// TIA Portal V20 export
FUNCTION_BLOCK "PR_MultiPosShuttle_Soft2.0 1_workflow_268c4d"   // FB49, LAD
{ S7_Optimized_Access := 'TRUE' }
// stored: MemoryReserve 100, SetENOAutomatically false
   VAR_INPUT
      iAutoRunning : Bool;
      iFaultReset : Bool;
      iGantry2Safe : Bool;
      iGantry_2Safe : Bool;
      iHIPOTTesSafe : Bool;
      iHIPOTTestOver : Bool;
      iHipotTestSafe : Bool;
      iInfeedGantrySafe : Bool;
      iOTS_Frm_Gantry : Bool;
      iPartPresent : Bool;
      iPartPrsent : Bool;
      iRTR_Frm_Gantry2 : Bool;
      iReset_fault : Bool;
      iShuttleAtGantry2Pos : Bool;
      iShuttleAtGantry_2Pos : Bool;
      iShuttleAtHIPOTPos : Bool;
      iShuttleAtHIPOTTestPos : Bool;
      iShuttleAtPartLoadPos : Bool;
      iSstMode : Bool;
      iSstPB : Bool;
   END_VAR
   VAR_OUTPUT
      qError : Array[0..10] of Bool;
      qHiPotTestStartCmd : Bool;
      qMessage : Array[0..10] of Bool;
      qRTR_To_InfeedGantry : Bool;
      qShuttleGantry_2PosCmd : Bool;
      qShuttleHIPOTTestPosCmd : Bool;
      qStateNo : Int;
      qShuttleReceivePosCmd : Bool;
   END_VAR
   VAR
      c10_ChkRecCond_T1 : Bool;
      c10_ChkRecCond_T2 : Bool;
      c10_ChkRecCond_T3 : Bool;
      c10_ChkRecCond_T4 : Bool;
      c10_ChkRecCond_T5 : Bool;
      c150_ChkOprnSts_T1 : Bool;
      c150_ChkOprnSts_T2 : Bool;
      c30_ChkPartPrsnt_T1 : Bool;
      c30_ChkPartPrsnt_T2 : Bool;
      s100_WtHipotTestOver : Bool;
      s100_WtHipotTestOver_T1 : Bool;
      s10_ChkRecCond : Bool;
      s10_ChkRecCond_T1 : Bool;
      s10_ChkRecCond_T2 : Bool;
      s10_ChkRecCond_T3 : Bool;
      s10_ChkRecCond_T4 : Bool;
      s10_ChkRecCond_T5 : Bool;
      s110_WtGantry2Safe : Bool;
      s110_WtGantry2Safe_T1 : Bool;
      s120_WtShtlGantry2Pos : Bool;
      s120_WtShtlGantry2Pos_T1 : Bool;
      s130_WtRTRFrmGantry2 : Bool;
      s130_WtRTRFrmGantry2_T1 : Bool;
      s140_WtPartAbsntGantry2Safe : Bool;
      s140_WtPartAbsntGantry2Safe_T1 : Bool;
      s150_ChkOprnSts : Bool;
      s150_ChkOprnSts_T1 : Bool;
      s150_ChkOprnSts_T2 : Bool;
      s1_WtResetRel : Bool;
      s1_WtResetRel_T1 : Bool;
      s20_WtFaultReset : Bool;
      s20_WtFaultReset_T1 : Bool;
      s30_ChkPartPrsnt : Bool;
      s30_ChkPartPrsnt_T1 : Bool;
      s30_ChkPartPrsnt_T2 : Bool;
      s40_WtAllSysSafe : Bool;
      s40_WtAllSysSafe_T1 : Bool;
      s50_WtShtlPartRcvPos : Bool;
      s50_WtShtlPartRcvPos_T1 : Bool;
      s60_WtOTSFrmGantry : Bool;
      s60_WtOTSFrmGantry_T1 : Bool;
      s70_WtPartPlcdGantrySafe : Bool;
      s70_WtPartPlcdGantrySafe_T1 : Bool;
      s80_WtHIPOTSafe : Bool;
      s80_WtHIPOTSafe_T1 : Bool;
      s90_WtShtlHIPOTPos : Bool;
      s90_WtShtlHIPOTPos_T1 : Bool;
      sHIPOTOprnOver : Bool;
      sHipotTestInProgress : Bool;
      sPickInProgress : Bool;
      sPlaceInProgress : Bool;
      sSst : Bool;
      sSstPulse : Bool;
      sSstRise : Bool;
      sStWtResetRel : Bool;
      sStWtResetRel_T1 : Bool;
   END_VAR
   VAR_TEMP
      tOne : Bool;
   END_VAR
   VAR_TEMP   // added for the SCL form of the ladder/FBD networks
      _w1 : Bool;
      _w2 : Bool;
      _w3 : Bool;
      _w4 : Bool;
   END_VAR
BEGIN

REGION Network 1
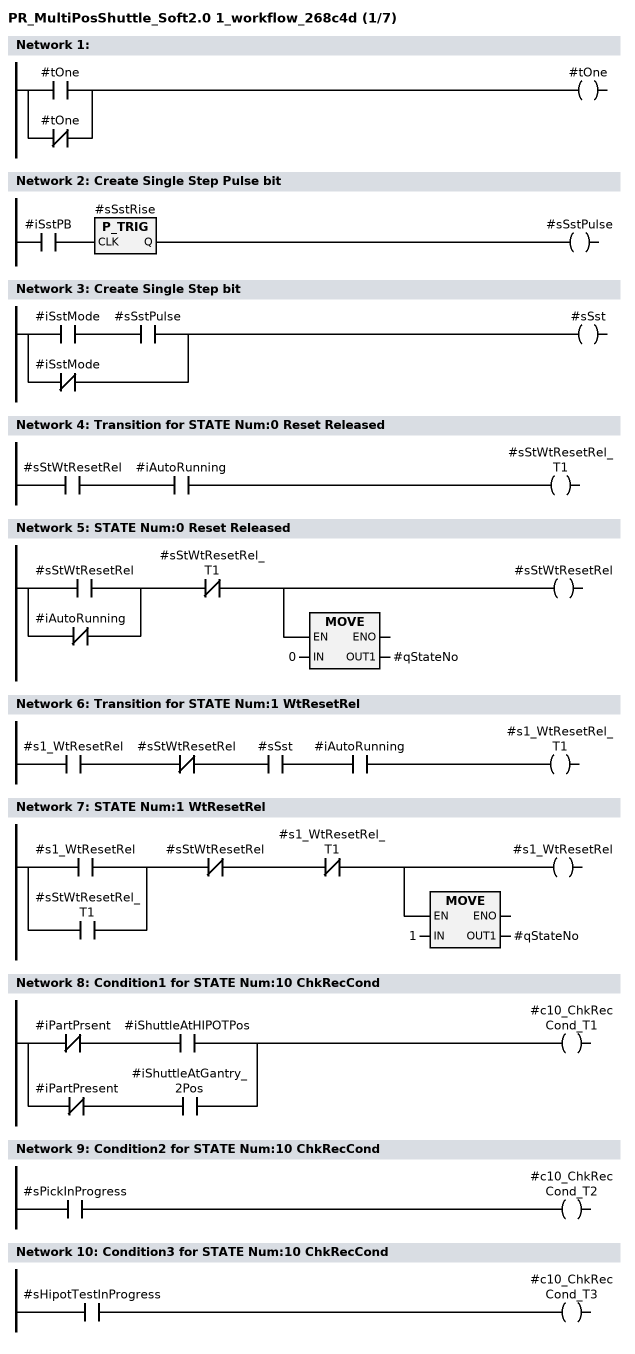
   RUNG wire#powerrail
      Contact( #tOne )
      wire#w1
      Coil( #tOne )
   END_RUNG
   RUNG wire#powerrail
      I_Contact( #tOne )
   END_RUNG wire#w1
   // the same network as SCL:
   #tOne := #tOne OR NOT #tOne;
END_REGION

REGION Network 2: Create Single Step Pulse bit
   RUNG wire#powerrail
      Contact( #iSstPB )
      P_Trig( #sSstRise )
      Coil( #sSstPulse )
   END_RUNG
   // the same network as SCL:
   #_w1 := #iSstPB AND NOT #sSstRise;   // rising edge
   #sSstRise := #iSstPB;
   #sSstPulse := #_w1;
END_REGION

REGION Network 3: Create Single Step bit
   RUNG wire#powerrail
      Contact( #iSstMode )
      Contact( #sSstPulse )
      wire#w1
      Coil( #sSst )
   END_RUNG
   RUNG wire#powerrail
      I_Contact( #iSstMode )
   END_RUNG wire#w1
   // the same network as SCL:
   #sSst := (#iSstMode AND #sSstPulse) OR NOT #iSstMode;
END_REGION

REGION Network 4: Transition for STATE Num:0 Reset Released
   RUNG wire#powerrail
      Contact( #sStWtResetRel )
      Contact( #iAutoRunning )
      Coil( #sStWtResetRel_T1 )
   END_RUNG
   // the same network as SCL:
   #sStWtResetRel_T1 := #sStWtResetRel AND #iAutoRunning;
END_REGION

REGION Network 5: STATE Num:0 Reset Released
   RUNG wire#powerrail
      Contact( #sStWtResetRel )
      wire#w1
      I_Contact( #sStWtResetRel_T1 )
      wire#w2
      Coil( #sStWtResetRel )
   END_RUNG
   RUNG wire#powerrail
      I_Contact( #iAutoRunning )
   END_RUNG wire#w1
   RUNG wire#w2
      { S7_GenerateENO := "TRUE" } Move(in := 0, out1 => #qStateNo)
   END_RUNG
   // the same network as SCL:
   #sStWtResetRel := (#sStWtResetRel OR NOT #iAutoRunning) AND NOT #sStWtResetRel_T1;
   IF #sStWtResetRel THEN #qStateNo := 0; END_IF;
END_REGION

REGION Network 6: Transition for STATE Num:1 WtResetRel
   RUNG wire#powerrail
      Contact( #s1_WtResetRel )
      I_Contact( #sStWtResetRel )
      Contact( #sSst )
      Contact( #iAutoRunning )
      Coil( #s1_WtResetRel_T1 )
   END_RUNG
   // the same network as SCL:
   #s1_WtResetRel_T1 := #s1_WtResetRel AND NOT #sStWtResetRel AND #sSst AND #iAutoRunning;
END_REGION

REGION Network 7: STATE Num:1 WtResetRel
   RUNG wire#powerrail
      Contact( #s1_WtResetRel )
      wire#w1
      I_Contact( #sStWtResetRel )
      I_Contact( #s1_WtResetRel_T1 )
      wire#w2
      Coil( #s1_WtResetRel )
   END_RUNG
   RUNG wire#powerrail
      Contact( #sStWtResetRel_T1 )
   END_RUNG wire#w1
   RUNG wire#w2
      { S7_GenerateENO := "TRUE" } Move(in := 1, out1 => #qStateNo)
   END_RUNG
   // the same network as SCL:
   #s1_WtResetRel := (#s1_WtResetRel OR #sStWtResetRel_T1) AND NOT #sStWtResetRel AND NOT #s1_WtResetRel_T1;
   IF #s1_WtResetRel THEN #qStateNo := 1; END_IF;
END_REGION

REGION Network 8: Condition1 for STATE Num:10 ChkRecCond
   RUNG wire#powerrail
      I_Contact( #iPartPrsent )
      Contact( #iShuttleAtHIPOTPos )
      wire#w1
      Coil( #c10_ChkRecCond_T1 )
   END_RUNG
   RUNG wire#powerrail
      I_Contact( #iPartPresent )
      Contact( #iShuttleAtGantry_2Pos )
   END_RUNG wire#w1
   // the same network as SCL:
   #c10_ChkRecCond_T1 := (NOT #iPartPrsent AND #iShuttleAtHIPOTPos) OR (NOT #iPartPresent AND #iShuttleAtGantry_2Pos);
END_REGION

REGION Network 9: Condition2 for STATE Num:10 ChkRecCond
   RUNG wire#powerrail
      Contact( #sPickInProgress )
      Coil( #c10_ChkRecCond_T2 )
   END_RUNG
   // the same network as SCL:
   #c10_ChkRecCond_T2 := #sPickInProgress;
END_REGION

REGION Network 10: Condition3 for STATE Num:10 ChkRecCond
   RUNG wire#powerrail
      Contact( #sHipotTestInProgress )
      Coil( #c10_ChkRecCond_T3 )
   END_RUNG
   // the same network as SCL:
   #c10_ChkRecCond_T3 := #sHipotTestInProgress;
END_REGION

REGION Network 11: Condition4 for STATE Num:10 ChkRecCond
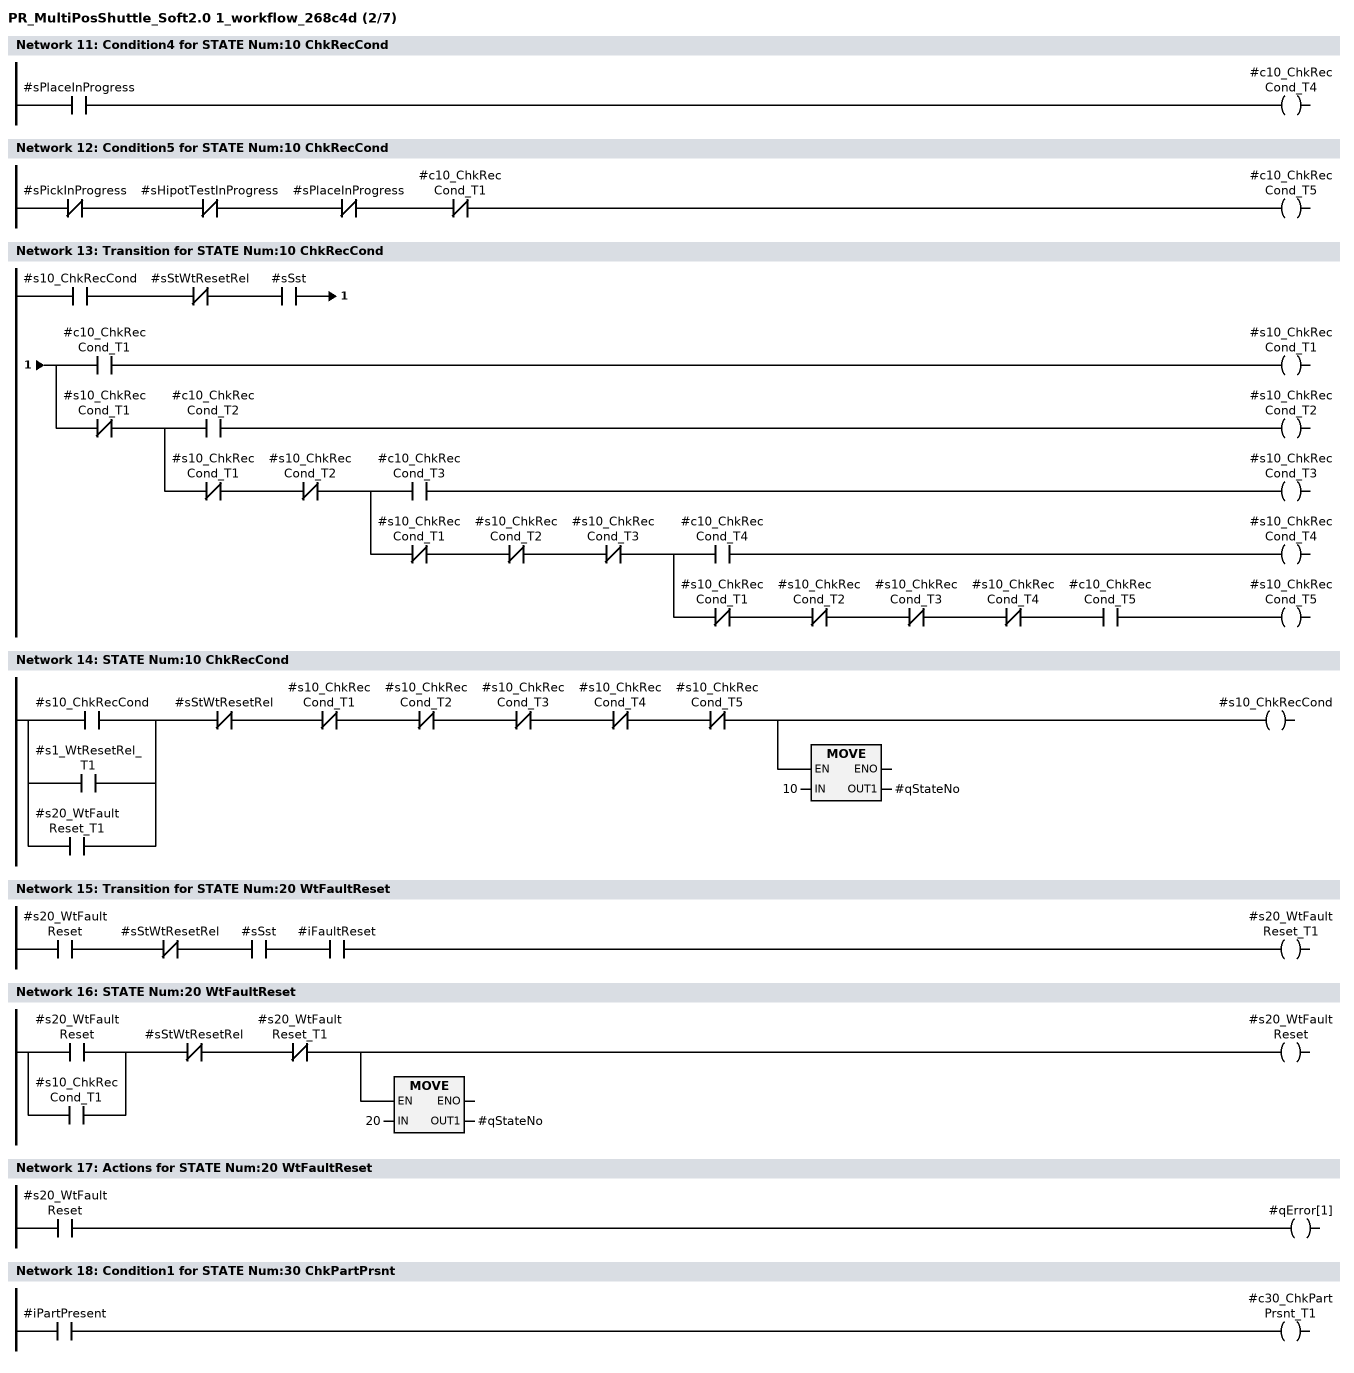
   RUNG wire#powerrail
      Contact( #sPlaceInProgress )
      Coil( #c10_ChkRecCond_T4 )
   END_RUNG
   // the same network as SCL:
   #c10_ChkRecCond_T4 := #sPlaceInProgress;
END_REGION

REGION Network 12: Condition5 for STATE Num:10 ChkRecCond
   RUNG wire#powerrail
      I_Contact( #sPickInProgress )
      I_Contact( #sHipotTestInProgress )
      I_Contact( #sPlaceInProgress )
      I_Contact( #c10_ChkRecCond_T1 )
      Coil( #c10_ChkRecCond_T5 )
   END_RUNG
   // the same network as SCL:
   #c10_ChkRecCond_T5 := NOT #sPickInProgress AND NOT #sHipotTestInProgress AND NOT #sPlaceInProgress AND NOT #c10_ChkRecCond_T1;
END_REGION

REGION Network 13: Transition for STATE Num:10 ChkRecCond
   RUNG wire#powerrail
      Contact( #s10_ChkRecCond )
      I_Contact( #sStWtResetRel )
      Contact( #sSst )
      wire#w1
      Contact( #c10_ChkRecCond_T1 )
      Coil( #s10_ChkRecCond_T1 )
   END_RUNG
   RUNG wire#w1
      I_Contact( #s10_ChkRecCond_T1 )
      wire#w2
      Contact( #c10_ChkRecCond_T2 )
      Coil( #s10_ChkRecCond_T2 )
   END_RUNG
   RUNG wire#w2
      I_Contact( #s10_ChkRecCond_T1 )
      I_Contact( #s10_ChkRecCond_T2 )
      wire#w3
      Contact( #c10_ChkRecCond_T3 )
      Coil( #s10_ChkRecCond_T3 )
   END_RUNG
   RUNG wire#w3
      I_Contact( #s10_ChkRecCond_T1 )
      I_Contact( #s10_ChkRecCond_T2 )
      I_Contact( #s10_ChkRecCond_T3 )
      wire#w4
      Contact( #c10_ChkRecCond_T4 )
      Coil( #s10_ChkRecCond_T4 )
   END_RUNG
   RUNG wire#w4
      I_Contact( #s10_ChkRecCond_T1 )
      I_Contact( #s10_ChkRecCond_T2 )
      I_Contact( #s10_ChkRecCond_T3 )
      I_Contact( #s10_ChkRecCond_T4 )
      Contact( #c10_ChkRecCond_T5 )
      Coil( #s10_ChkRecCond_T5 )
   END_RUNG
   // the same network as SCL:
   #_w1 := #s10_ChkRecCond AND NOT #sStWtResetRel AND #sSst;
   #s10_ChkRecCond_T1 := #_w1 AND #c10_ChkRecCond_T1;
   #_w2 := #_w1 AND NOT #s10_ChkRecCond_T1;
   #s10_ChkRecCond_T2 := #_w2 AND #c10_ChkRecCond_T2;
   #_w3 := #_w2 AND NOT #s10_ChkRecCond_T1 AND NOT #s10_ChkRecCond_T2;
   #s10_ChkRecCond_T3 := #_w3 AND #c10_ChkRecCond_T3;
   #_w4 := #_w3 AND NOT #s10_ChkRecCond_T1 AND NOT #s10_ChkRecCond_T2 AND NOT #s10_ChkRecCond_T3;
   #s10_ChkRecCond_T4 := #_w4 AND #c10_ChkRecCond_T4;
   #s10_ChkRecCond_T5 := #_w4 AND NOT #s10_ChkRecCond_T1 AND NOT #s10_ChkRecCond_T2 AND NOT #s10_ChkRecCond_T3 AND NOT #s10_ChkRecCond_T4 AND #c10_ChkRecCond_T5;
END_REGION

REGION Network 14: STATE Num:10 ChkRecCond
   RUNG wire#powerrail
      Contact( #s10_ChkRecCond )
      wire#w1
      I_Contact( #sStWtResetRel )
      I_Contact( #s10_ChkRecCond_T1 )
      I_Contact( #s10_ChkRecCond_T2 )
      I_Contact( #s10_ChkRecCond_T3 )
      I_Contact( #s10_ChkRecCond_T4 )
      I_Contact( #s10_ChkRecCond_T5 )
      wire#w2
      Coil( #s10_ChkRecCond )
   END_RUNG
   RUNG wire#powerrail
      Contact( #s1_WtResetRel_T1 )
   END_RUNG wire#w1
   RUNG wire#powerrail
      Contact( #s20_WtFaultReset_T1 )
   END_RUNG wire#w1
   RUNG wire#w2
      { S7_GenerateENO := "TRUE" } Move(in := 10, out1 => #qStateNo)
   END_RUNG
   // the same network as SCL:
   #s10_ChkRecCond := (#s10_ChkRecCond OR #s1_WtResetRel_T1 OR #s20_WtFaultReset_T1) AND NOT #sStWtResetRel AND NOT #s10_ChkRecCond_T1 AND NOT #s10_ChkRecCond_T2 AND NOT #s10_ChkRecCond_T3 AND NOT #s10_ChkRecCond_T4 AND NOT #s10_ChkRecCond_T5;
   IF #s10_ChkRecCond THEN #qStateNo := 10; END_IF;
END_REGION

REGION Network 15: Transition for STATE Num:20 WtFaultReset
   RUNG wire#powerrail
      Contact( #s20_WtFaultReset )
      I_Contact( #sStWtResetRel )
      Contact( #sSst )
      Contact( #iFaultReset )
      Coil( #s20_WtFaultReset_T1 )
   END_RUNG
   // the same network as SCL:
   #s20_WtFaultReset_T1 := #s20_WtFaultReset AND NOT #sStWtResetRel AND #sSst AND #iFaultReset;
END_REGION

REGION Network 16: STATE Num:20 WtFaultReset
   RUNG wire#powerrail
      Contact( #s20_WtFaultReset )
      wire#w1
      I_Contact( #sStWtResetRel )
      I_Contact( #s20_WtFaultReset_T1 )
      wire#w2
      Coil( #s20_WtFaultReset )
   END_RUNG
   RUNG wire#powerrail
      Contact( #s10_ChkRecCond_T1 )
   END_RUNG wire#w1
   RUNG wire#w2
      { S7_GenerateENO := "TRUE" } Move(in := 20, out1 => #qStateNo)
   END_RUNG
   // the same network as SCL:
   #s20_WtFaultReset := (#s20_WtFaultReset OR #s10_ChkRecCond_T1) AND NOT #sStWtResetRel AND NOT #s20_WtFaultReset_T1;
   IF #s20_WtFaultReset THEN #qStateNo := 20; END_IF;
END_REGION

REGION Network 17: Actions for STATE Num:20 WtFaultReset
   RUNG wire#powerrail
      Contact( #s20_WtFaultReset )
      Coil( #qError[1] )
   END_RUNG
   // the same network as SCL:
   #qError[1] := #s20_WtFaultReset;
END_REGION

REGION Network 18: Condition1 for STATE Num:30 ChkPartPrsnt
   RUNG wire#powerrail
      Contact( #iPartPresent )
      Coil( #c30_ChkPartPrsnt_T1 )
   END_RUNG
   // the same network as SCL:
   #c30_ChkPartPrsnt_T1 := #iPartPresent;
END_REGION

REGION Network 19: Condition2 for STATE Num:30 ChkPartPrsnt
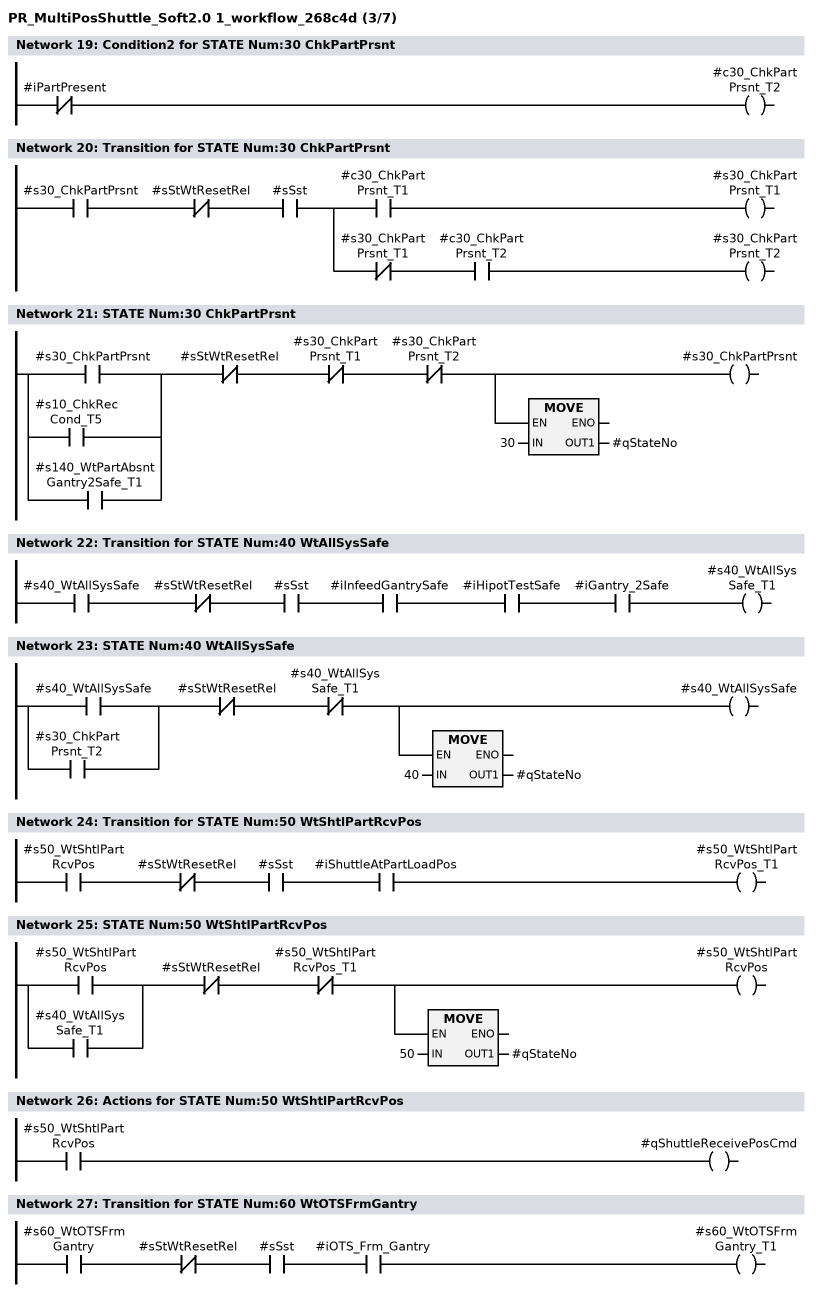
   RUNG wire#powerrail
      I_Contact( #iPartPresent )
      Coil( #c30_ChkPartPrsnt_T2 )
   END_RUNG
   // the same network as SCL:
   #c30_ChkPartPrsnt_T2 := NOT #iPartPresent;
END_REGION

REGION Network 20: Transition for STATE Num:30 ChkPartPrsnt
   RUNG wire#powerrail
      Contact( #s30_ChkPartPrsnt )
      I_Contact( #sStWtResetRel )
      Contact( #sSst )
      wire#w1
      Contact( #c30_ChkPartPrsnt_T1 )
      Coil( #s30_ChkPartPrsnt_T1 )
   END_RUNG
   RUNG wire#w1
      I_Contact( #s30_ChkPartPrsnt_T1 )
      Contact( #c30_ChkPartPrsnt_T2 )
      Coil( #s30_ChkPartPrsnt_T2 )
   END_RUNG
   // the same network as SCL:
   #_w1 := #s30_ChkPartPrsnt AND NOT #sStWtResetRel AND #sSst;
   #s30_ChkPartPrsnt_T1 := #_w1 AND #c30_ChkPartPrsnt_T1;
   #s30_ChkPartPrsnt_T2 := #_w1 AND NOT #s30_ChkPartPrsnt_T1 AND #c30_ChkPartPrsnt_T2;
END_REGION

REGION Network 21: STATE Num:30 ChkPartPrsnt
   RUNG wire#powerrail
      Contact( #s30_ChkPartPrsnt )
      wire#w1
      I_Contact( #sStWtResetRel )
      I_Contact( #s30_ChkPartPrsnt_T1 )
      I_Contact( #s30_ChkPartPrsnt_T2 )
      wire#w2
      Coil( #s30_ChkPartPrsnt )
   END_RUNG
   RUNG wire#powerrail
      Contact( #s10_ChkRecCond_T5 )
   END_RUNG wire#w1
   RUNG wire#powerrail
      Contact( #s140_WtPartAbsntGantry2Safe_T1 )
   END_RUNG wire#w1
   RUNG wire#w2
      { S7_GenerateENO := "TRUE" } Move(in := 30, out1 => #qStateNo)
   END_RUNG
   // the same network as SCL:
   #s30_ChkPartPrsnt := (#s30_ChkPartPrsnt OR #s10_ChkRecCond_T5 OR #s140_WtPartAbsntGantry2Safe_T1) AND NOT #sStWtResetRel AND NOT #s30_ChkPartPrsnt_T1 AND NOT #s30_ChkPartPrsnt_T2;
   IF #s30_ChkPartPrsnt THEN #qStateNo := 30; END_IF;
END_REGION

REGION Network 22: Transition for STATE Num:40 WtAllSysSafe
   RUNG wire#powerrail
      Contact( #s40_WtAllSysSafe )
      I_Contact( #sStWtResetRel )
      Contact( #sSst )
      Contact( #iInfeedGantrySafe )
      Contact( #iHipotTestSafe )
      Contact( #iGantry_2Safe )
      Coil( #s40_WtAllSysSafe_T1 )
   END_RUNG
   // the same network as SCL:
   #s40_WtAllSysSafe_T1 := #s40_WtAllSysSafe AND NOT #sStWtResetRel AND #sSst AND #iInfeedGantrySafe AND #iHipotTestSafe AND #iGantry_2Safe;
END_REGION

REGION Network 23: STATE Num:40 WtAllSysSafe
   RUNG wire#powerrail
      Contact( #s40_WtAllSysSafe )
      wire#w1
      I_Contact( #sStWtResetRel )
      I_Contact( #s40_WtAllSysSafe_T1 )
      wire#w2
      Coil( #s40_WtAllSysSafe )
   END_RUNG
   RUNG wire#powerrail
      Contact( #s30_ChkPartPrsnt_T2 )
   END_RUNG wire#w1
   RUNG wire#w2
      { S7_GenerateENO := "TRUE" } Move(in := 40, out1 => #qStateNo)
   END_RUNG
   // the same network as SCL:
   #s40_WtAllSysSafe := (#s40_WtAllSysSafe OR #s30_ChkPartPrsnt_T2) AND NOT #sStWtResetRel AND NOT #s40_WtAllSysSafe_T1;
   IF #s40_WtAllSysSafe THEN #qStateNo := 40; END_IF;
END_REGION

REGION Network 24: Transition for STATE Num:50 WtShtlPartRcvPos
   RUNG wire#powerrail
      Contact( #s50_WtShtlPartRcvPos )
      I_Contact( #sStWtResetRel )
      Contact( #sSst )
      Contact( #iShuttleAtPartLoadPos )
      Coil( #s50_WtShtlPartRcvPos_T1 )
   END_RUNG
   // the same network as SCL:
   #s50_WtShtlPartRcvPos_T1 := #s50_WtShtlPartRcvPos AND NOT #sStWtResetRel AND #sSst AND #iShuttleAtPartLoadPos;
END_REGION

REGION Network 25: STATE Num:50 WtShtlPartRcvPos
   RUNG wire#powerrail
      Contact( #s50_WtShtlPartRcvPos )
      wire#w1
      I_Contact( #sStWtResetRel )
      I_Contact( #s50_WtShtlPartRcvPos_T1 )
      wire#w2
      Coil( #s50_WtShtlPartRcvPos )
   END_RUNG
   RUNG wire#powerrail
      Contact( #s40_WtAllSysSafe_T1 )
   END_RUNG wire#w1
   RUNG wire#w2
      { S7_GenerateENO := "TRUE" } Move(in := 50, out1 => #qStateNo)
   END_RUNG
   // the same network as SCL:
   #s50_WtShtlPartRcvPos := (#s50_WtShtlPartRcvPos OR #s40_WtAllSysSafe_T1) AND NOT #sStWtResetRel AND NOT #s50_WtShtlPartRcvPos_T1;
   IF #s50_WtShtlPartRcvPos THEN #qStateNo := 50; END_IF;
END_REGION

REGION Network 26: Actions for STATE Num:50 WtShtlPartRcvPos
   RUNG wire#powerrail
      Contact( #s50_WtShtlPartRcvPos )
      Coil( #qShuttleReceivePosCmd )
   END_RUNG
   // the same network as SCL:
   #qShuttleReceivePosCmd := #s50_WtShtlPartRcvPos;
END_REGION

REGION Network 27: Transition for STATE Num:60 WtOTSFrmGantry
   RUNG wire#powerrail
      Contact( #s60_WtOTSFrmGantry )
      I_Contact( #sStWtResetRel )
      Contact( #sSst )
      Contact( #iOTS_Frm_Gantry )
      Coil( #s60_WtOTSFrmGantry_T1 )
   END_RUNG
   // the same network as SCL:
   #s60_WtOTSFrmGantry_T1 := #s60_WtOTSFrmGantry AND NOT #sStWtResetRel AND #sSst AND #iOTS_Frm_Gantry;
END_REGION

REGION Network 28: STATE Num:60 WtOTSFrmGantry
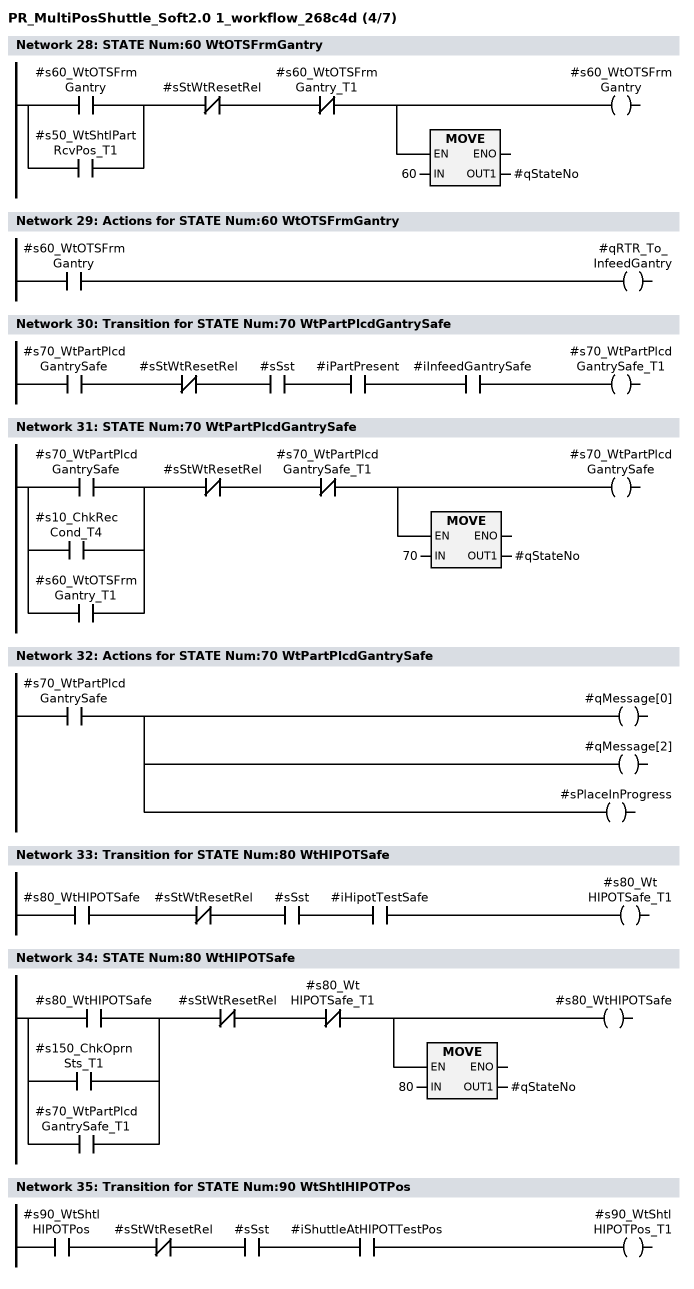
   RUNG wire#powerrail
      Contact( #s60_WtOTSFrmGantry )
      wire#w1
      I_Contact( #sStWtResetRel )
      I_Contact( #s60_WtOTSFrmGantry_T1 )
      wire#w2
      Coil( #s60_WtOTSFrmGantry )
   END_RUNG
   RUNG wire#powerrail
      Contact( #s50_WtShtlPartRcvPos_T1 )
   END_RUNG wire#w1
   RUNG wire#w2
      { S7_GenerateENO := "TRUE" } Move(in := 60, out1 => #qStateNo)
   END_RUNG
   // the same network as SCL:
   #s60_WtOTSFrmGantry := (#s60_WtOTSFrmGantry OR #s50_WtShtlPartRcvPos_T1) AND NOT #sStWtResetRel AND NOT #s60_WtOTSFrmGantry_T1;
   IF #s60_WtOTSFrmGantry THEN #qStateNo := 60; END_IF;
END_REGION

REGION Network 29: Actions for STATE Num:60 WtOTSFrmGantry
   RUNG wire#powerrail
      Contact( #s60_WtOTSFrmGantry )
      Coil( #qRTR_To_InfeedGantry )
   END_RUNG
   // the same network as SCL:
   #qRTR_To_InfeedGantry := #s60_WtOTSFrmGantry;
END_REGION

REGION Network 30: Transition for STATE Num:70 WtPartPlcdGantrySafe
   RUNG wire#powerrail
      Contact( #s70_WtPartPlcdGantrySafe )
      I_Contact( #sStWtResetRel )
      Contact( #sSst )
      Contact( #iPartPresent )
      Contact( #iInfeedGantrySafe )
      Coil( #s70_WtPartPlcdGantrySafe_T1 )
   END_RUNG
   // the same network as SCL:
   #s70_WtPartPlcdGantrySafe_T1 := #s70_WtPartPlcdGantrySafe AND NOT #sStWtResetRel AND #sSst AND #iPartPresent AND #iInfeedGantrySafe;
END_REGION

REGION Network 31: STATE Num:70 WtPartPlcdGantrySafe
   RUNG wire#powerrail
      Contact( #s70_WtPartPlcdGantrySafe )
      wire#w1
      I_Contact( #sStWtResetRel )
      I_Contact( #s70_WtPartPlcdGantrySafe_T1 )
      wire#w2
      Coil( #s70_WtPartPlcdGantrySafe )
   END_RUNG
   RUNG wire#powerrail
      Contact( #s10_ChkRecCond_T4 )
   END_RUNG wire#w1
   RUNG wire#powerrail
      Contact( #s60_WtOTSFrmGantry_T1 )
   END_RUNG wire#w1
   RUNG wire#w2
      { S7_GenerateENO := "TRUE" } Move(in := 70, out1 => #qStateNo)
   END_RUNG
   // the same network as SCL:
   #s70_WtPartPlcdGantrySafe := (#s70_WtPartPlcdGantrySafe OR #s10_ChkRecCond_T4 OR #s60_WtOTSFrmGantry_T1) AND NOT #sStWtResetRel AND NOT #s70_WtPartPlcdGantrySafe_T1;
   IF #s70_WtPartPlcdGantrySafe THEN #qStateNo := 70; END_IF;
END_REGION

REGION Network 32: Actions for STATE Num:70 WtPartPlcdGantrySafe
   RUNG wire#powerrail
      Contact( #s70_WtPartPlcdGantrySafe )
      wire#w1
      Coil( #qMessage[0] )
   END_RUNG
   RUNG wire#w1
      Coil( #qMessage[2] )
   END_RUNG
   RUNG wire#w1
      Coil( #sPlaceInProgress )
   END_RUNG
   // the same network as SCL:
   #qMessage[0] := #s70_WtPartPlcdGantrySafe;
   #qMessage[2] := #s70_WtPartPlcdGantrySafe;
   #sPlaceInProgress := #s70_WtPartPlcdGantrySafe;
END_REGION

REGION Network 33: Transition for STATE Num:80 WtHIPOTSafe
   RUNG wire#powerrail
      Contact( #s80_WtHIPOTSafe )
      I_Contact( #sStWtResetRel )
      Contact( #sSst )
      Contact( #iHipotTestSafe )
      Coil( #s80_WtHIPOTSafe_T1 )
   END_RUNG
   // the same network as SCL:
   #s80_WtHIPOTSafe_T1 := #s80_WtHIPOTSafe AND NOT #sStWtResetRel AND #sSst AND #iHipotTestSafe;
END_REGION

REGION Network 34: STATE Num:80 WtHIPOTSafe
   RUNG wire#powerrail
      Contact( #s80_WtHIPOTSafe )
      wire#w1
      I_Contact( #sStWtResetRel )
      I_Contact( #s80_WtHIPOTSafe_T1 )
      wire#w2
      Coil( #s80_WtHIPOTSafe )
   END_RUNG
   RUNG wire#powerrail
      Contact( #s150_ChkOprnSts_T1 )
   END_RUNG wire#w1
   RUNG wire#powerrail
      Contact( #s70_WtPartPlcdGantrySafe_T1 )
   END_RUNG wire#w1
   RUNG wire#w2
      { S7_GenerateENO := "TRUE" } Move(in := 80, out1 => #qStateNo)
   END_RUNG
   // the same network as SCL:
   #s80_WtHIPOTSafe := (#s80_WtHIPOTSafe OR #s150_ChkOprnSts_T1 OR #s70_WtPartPlcdGantrySafe_T1) AND NOT #sStWtResetRel AND NOT #s80_WtHIPOTSafe_T1;
   IF #s80_WtHIPOTSafe THEN #qStateNo := 80; END_IF;
END_REGION

REGION Network 35: Transition for STATE Num:90 WtShtlHIPOTPos
   RUNG wire#powerrail
      Contact( #s90_WtShtlHIPOTPos )
      I_Contact( #sStWtResetRel )
      Contact( #sSst )
      Contact( #iShuttleAtHIPOTTestPos )
      Coil( #s90_WtShtlHIPOTPos_T1 )
   END_RUNG
   // the same network as SCL:
   #s90_WtShtlHIPOTPos_T1 := #s90_WtShtlHIPOTPos AND NOT #sStWtResetRel AND #sSst AND #iShuttleAtHIPOTTestPos;
END_REGION

REGION Network 36: STATE Num:90 WtShtlHIPOTPos
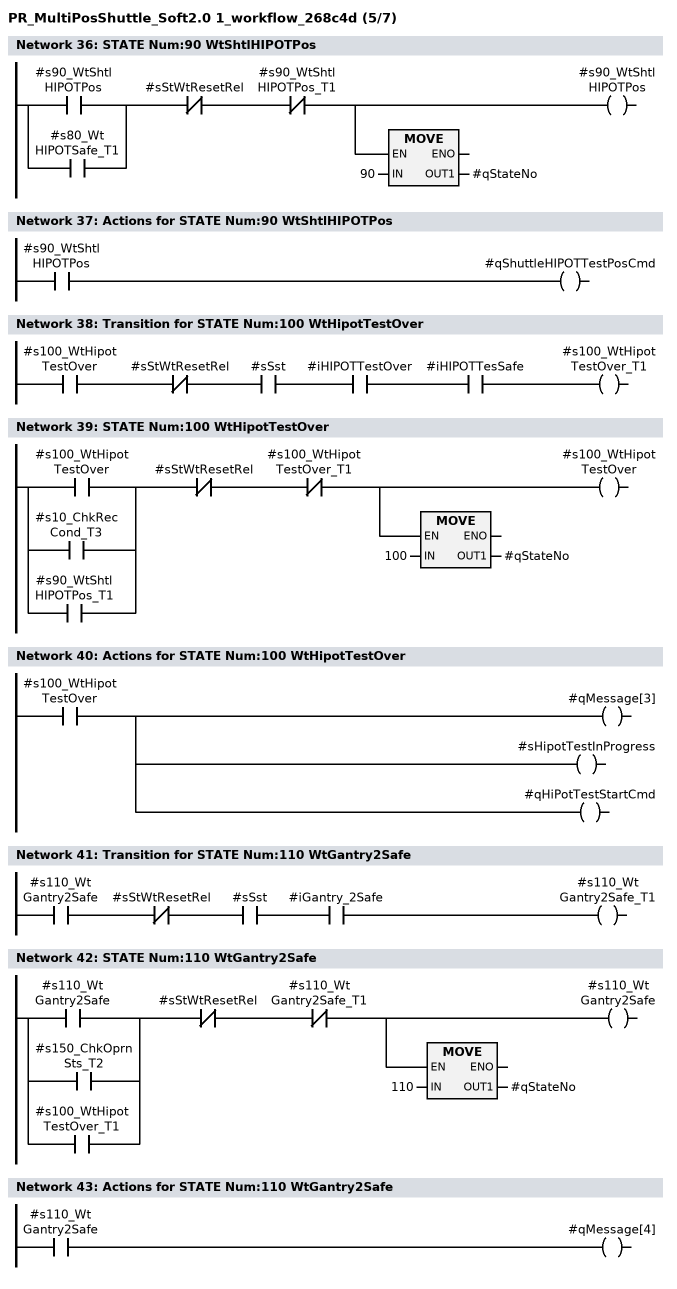
   RUNG wire#powerrail
      Contact( #s90_WtShtlHIPOTPos )
      wire#w1
      I_Contact( #sStWtResetRel )
      I_Contact( #s90_WtShtlHIPOTPos_T1 )
      wire#w2
      Coil( #s90_WtShtlHIPOTPos )
   END_RUNG
   RUNG wire#powerrail
      Contact( #s80_WtHIPOTSafe_T1 )
   END_RUNG wire#w1
   RUNG wire#w2
      { S7_GenerateENO := "TRUE" } Move(in := 90, out1 => #qStateNo)
   END_RUNG
   // the same network as SCL:
   #s90_WtShtlHIPOTPos := (#s90_WtShtlHIPOTPos OR #s80_WtHIPOTSafe_T1) AND NOT #sStWtResetRel AND NOT #s90_WtShtlHIPOTPos_T1;
   IF #s90_WtShtlHIPOTPos THEN #qStateNo := 90; END_IF;
END_REGION

REGION Network 37: Actions for STATE Num:90 WtShtlHIPOTPos
   RUNG wire#powerrail
      Contact( #s90_WtShtlHIPOTPos )
      Coil( #qShuttleHIPOTTestPosCmd )
   END_RUNG
   // the same network as SCL:
   #qShuttleHIPOTTestPosCmd := #s90_WtShtlHIPOTPos;
END_REGION

REGION Network 38: Transition for STATE Num:100 WtHipotTestOver
   RUNG wire#powerrail
      Contact( #s100_WtHipotTestOver )
      I_Contact( #sStWtResetRel )
      Contact( #sSst )
      Contact( #iHIPOTTestOver )
      Contact( #iHIPOTTesSafe )
      Coil( #s100_WtHipotTestOver_T1 )
   END_RUNG
   // the same network as SCL:
   #s100_WtHipotTestOver_T1 := #s100_WtHipotTestOver AND NOT #sStWtResetRel AND #sSst AND #iHIPOTTestOver AND #iHIPOTTesSafe;
END_REGION

REGION Network 39: STATE Num:100 WtHipotTestOver
   RUNG wire#powerrail
      Contact( #s100_WtHipotTestOver )
      wire#w1
      I_Contact( #sStWtResetRel )
      I_Contact( #s100_WtHipotTestOver_T1 )
      wire#w2
      Coil( #s100_WtHipotTestOver )
   END_RUNG
   RUNG wire#powerrail
      Contact( #s10_ChkRecCond_T3 )
   END_RUNG wire#w1
   RUNG wire#powerrail
      Contact( #s90_WtShtlHIPOTPos_T1 )
   END_RUNG wire#w1
   RUNG wire#w2
      { S7_GenerateENO := "TRUE" } Move(in := 100, out1 => #qStateNo)
   END_RUNG
   // the same network as SCL:
   #s100_WtHipotTestOver := (#s100_WtHipotTestOver OR #s10_ChkRecCond_T3 OR #s90_WtShtlHIPOTPos_T1) AND NOT #sStWtResetRel AND NOT #s100_WtHipotTestOver_T1;
   IF #s100_WtHipotTestOver THEN #qStateNo := 100; END_IF;
END_REGION

REGION Network 40: Actions for STATE Num:100 WtHipotTestOver
   RUNG wire#powerrail
      Contact( #s100_WtHipotTestOver )
      wire#w1
      Coil( #qMessage[3] )
   END_RUNG
   RUNG wire#w1
      Coil( #sHipotTestInProgress )
   END_RUNG
   RUNG wire#w1
      Coil( #qHiPotTestStartCmd )
   END_RUNG
   // the same network as SCL:
   #qMessage[3] := #s100_WtHipotTestOver;
   #sHipotTestInProgress := #s100_WtHipotTestOver;
   #qHiPotTestStartCmd := #s100_WtHipotTestOver;
END_REGION

REGION Network 41: Transition for STATE Num:110 WtGantry2Safe
   RUNG wire#powerrail
      Contact( #s110_WtGantry2Safe )
      I_Contact( #sStWtResetRel )
      Contact( #sSst )
      Contact( #iGantry_2Safe )
      Coil( #s110_WtGantry2Safe_T1 )
   END_RUNG
   // the same network as SCL:
   #s110_WtGantry2Safe_T1 := #s110_WtGantry2Safe AND NOT #sStWtResetRel AND #sSst AND #iGantry_2Safe;
END_REGION

REGION Network 42: STATE Num:110 WtGantry2Safe
   RUNG wire#powerrail
      Contact( #s110_WtGantry2Safe )
      wire#w1
      I_Contact( #sStWtResetRel )
      I_Contact( #s110_WtGantry2Safe_T1 )
      wire#w2
      Coil( #s110_WtGantry2Safe )
   END_RUNG
   RUNG wire#powerrail
      Contact( #s150_ChkOprnSts_T2 )
   END_RUNG wire#w1
   RUNG wire#powerrail
      Contact( #s100_WtHipotTestOver_T1 )
   END_RUNG wire#w1
   RUNG wire#w2
      { S7_GenerateENO := "TRUE" } Move(in := 110, out1 => #qStateNo)
   END_RUNG
   // the same network as SCL:
   #s110_WtGantry2Safe := (#s110_WtGantry2Safe OR #s150_ChkOprnSts_T2 OR #s100_WtHipotTestOver_T1) AND NOT #sStWtResetRel AND NOT #s110_WtGantry2Safe_T1;
   IF #s110_WtGantry2Safe THEN #qStateNo := 110; END_IF;
END_REGION

REGION Network 43: Actions for STATE Num:110 WtGantry2Safe
   RUNG wire#powerrail
      Contact( #s110_WtGantry2Safe )
      Coil( #qMessage[4] )
   END_RUNG
   // the same network as SCL:
   #qMessage[4] := #s110_WtGantry2Safe;
END_REGION

REGION Network 44: Transition for STATE Num:120 WtShtlGantry2Pos
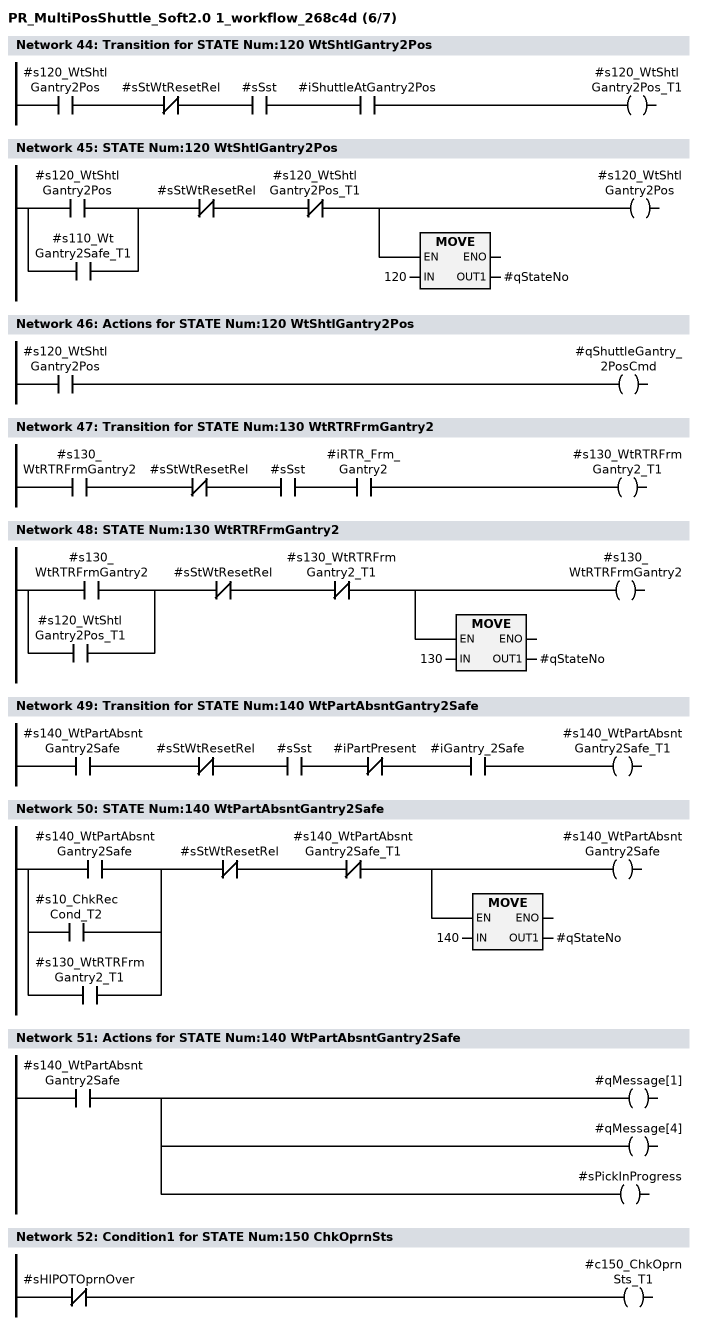
   RUNG wire#powerrail
      Contact( #s120_WtShtlGantry2Pos )
      I_Contact( #sStWtResetRel )
      Contact( #sSst )
      Contact( #iShuttleAtGantry2Pos )
      Coil( #s120_WtShtlGantry2Pos_T1 )
   END_RUNG
   // the same network as SCL:
   #s120_WtShtlGantry2Pos_T1 := #s120_WtShtlGantry2Pos AND NOT #sStWtResetRel AND #sSst AND #iShuttleAtGantry2Pos;
END_REGION

REGION Network 45: STATE Num:120 WtShtlGantry2Pos
   RUNG wire#powerrail
      Contact( #s120_WtShtlGantry2Pos )
      wire#w1
      I_Contact( #sStWtResetRel )
      I_Contact( #s120_WtShtlGantry2Pos_T1 )
      wire#w2
      Coil( #s120_WtShtlGantry2Pos )
   END_RUNG
   RUNG wire#powerrail
      Contact( #s110_WtGantry2Safe_T1 )
   END_RUNG wire#w1
   RUNG wire#w2
      { S7_GenerateENO := "TRUE" } Move(in := 120, out1 => #qStateNo)
   END_RUNG
   // the same network as SCL:
   #s120_WtShtlGantry2Pos := (#s120_WtShtlGantry2Pos OR #s110_WtGantry2Safe_T1) AND NOT #sStWtResetRel AND NOT #s120_WtShtlGantry2Pos_T1;
   IF #s120_WtShtlGantry2Pos THEN #qStateNo := 120; END_IF;
END_REGION

REGION Network 46: Actions for STATE Num:120 WtShtlGantry2Pos
   RUNG wire#powerrail
      Contact( #s120_WtShtlGantry2Pos )
      Coil( #qShuttleGantry_2PosCmd )
   END_RUNG
   // the same network as SCL:
   #qShuttleGantry_2PosCmd := #s120_WtShtlGantry2Pos;
END_REGION

REGION Network 47: Transition for STATE Num:130 WtRTRFrmGantry2
   RUNG wire#powerrail
      Contact( #s130_WtRTRFrmGantry2 )
      I_Contact( #sStWtResetRel )
      Contact( #sSst )
      Contact( #iRTR_Frm_Gantry2 )
      Coil( #s130_WtRTRFrmGantry2_T1 )
   END_RUNG
   // the same network as SCL:
   #s130_WtRTRFrmGantry2_T1 := #s130_WtRTRFrmGantry2 AND NOT #sStWtResetRel AND #sSst AND #iRTR_Frm_Gantry2;
END_REGION

REGION Network 48: STATE Num:130 WtRTRFrmGantry2
   RUNG wire#powerrail
      Contact( #s130_WtRTRFrmGantry2 )
      wire#w1
      I_Contact( #sStWtResetRel )
      I_Contact( #s130_WtRTRFrmGantry2_T1 )
      wire#w2
      Coil( #s130_WtRTRFrmGantry2 )
   END_RUNG
   RUNG wire#powerrail
      Contact( #s120_WtShtlGantry2Pos_T1 )
   END_RUNG wire#w1
   RUNG wire#w2
      { S7_GenerateENO := "TRUE" } Move(in := 130, out1 => #qStateNo)
   END_RUNG
   // the same network as SCL:
   #s130_WtRTRFrmGantry2 := (#s130_WtRTRFrmGantry2 OR #s120_WtShtlGantry2Pos_T1) AND NOT #sStWtResetRel AND NOT #s130_WtRTRFrmGantry2_T1;
   IF #s130_WtRTRFrmGantry2 THEN #qStateNo := 130; END_IF;
END_REGION

REGION Network 49: Transition for STATE Num:140 WtPartAbsntGantry2Safe
   RUNG wire#powerrail
      Contact( #s140_WtPartAbsntGantry2Safe )
      I_Contact( #sStWtResetRel )
      Contact( #sSst )
      I_Contact( #iPartPresent )
      Contact( #iGantry_2Safe )
      Coil( #s140_WtPartAbsntGantry2Safe_T1 )
   END_RUNG
   // the same network as SCL:
   #s140_WtPartAbsntGantry2Safe_T1 := #s140_WtPartAbsntGantry2Safe AND NOT #sStWtResetRel AND #sSst AND NOT #iPartPresent AND #iGantry_2Safe;
END_REGION

REGION Network 50: STATE Num:140 WtPartAbsntGantry2Safe
   RUNG wire#powerrail
      Contact( #s140_WtPartAbsntGantry2Safe )
      wire#w1
      I_Contact( #sStWtResetRel )
      I_Contact( #s140_WtPartAbsntGantry2Safe_T1 )
      wire#w2
      Coil( #s140_WtPartAbsntGantry2Safe )
   END_RUNG
   RUNG wire#powerrail
      Contact( #s10_ChkRecCond_T2 )
   END_RUNG wire#w1
   RUNG wire#powerrail
      Contact( #s130_WtRTRFrmGantry2_T1 )
   END_RUNG wire#w1
   RUNG wire#w2
      { S7_GenerateENO := "TRUE" } Move(in := 140, out1 => #qStateNo)
   END_RUNG
   // the same network as SCL:
   #s140_WtPartAbsntGantry2Safe := (#s140_WtPartAbsntGantry2Safe OR #s10_ChkRecCond_T2 OR #s130_WtRTRFrmGantry2_T1) AND NOT #sStWtResetRel AND NOT #s140_WtPartAbsntGantry2Safe_T1;
   IF #s140_WtPartAbsntGantry2Safe THEN #qStateNo := 140; END_IF;
END_REGION

REGION Network 51: Actions for STATE Num:140 WtPartAbsntGantry2Safe
   RUNG wire#powerrail
      Contact( #s140_WtPartAbsntGantry2Safe )
      wire#w1
      Coil( #qMessage[1] )
   END_RUNG
   RUNG wire#w1
      Coil( #qMessage[4] )
   END_RUNG
   RUNG wire#w1
      Coil( #sPickInProgress )
   END_RUNG
   // the same network as SCL:
   #qMessage[1] := #s140_WtPartAbsntGantry2Safe;
   #qMessage[4] := #s140_WtPartAbsntGantry2Safe;
   #sPickInProgress := #s140_WtPartAbsntGantry2Safe;
END_REGION

REGION Network 52: Condition1 for STATE Num:150 ChkOprnSts
   RUNG wire#powerrail
      I_Contact( #sHIPOTOprnOver )
      Coil( #c150_ChkOprnSts_T1 )
   END_RUNG
   // the same network as SCL:
   #c150_ChkOprnSts_T1 := NOT #sHIPOTOprnOver;
END_REGION

REGION Network 53: Condition2 for STATE Num:150 ChkOprnSts
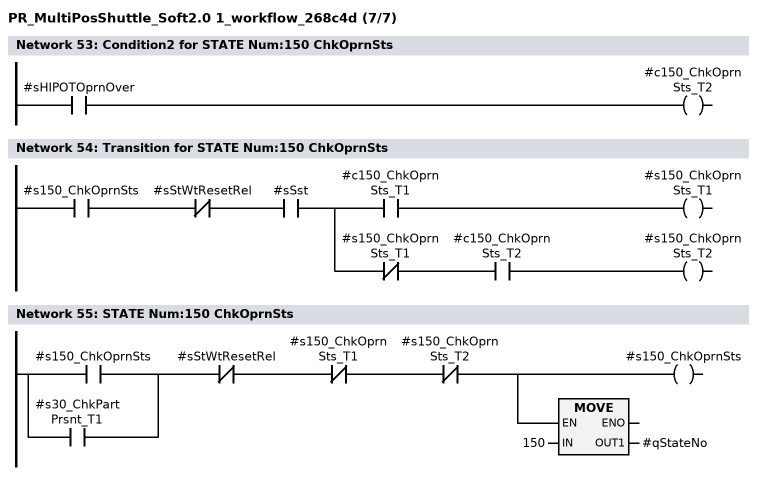
   RUNG wire#powerrail
      Contact( #sHIPOTOprnOver )
      Coil( #c150_ChkOprnSts_T2 )
   END_RUNG
   // the same network as SCL:
   #c150_ChkOprnSts_T2 := #sHIPOTOprnOver;
END_REGION

REGION Network 54: Transition for STATE Num:150 ChkOprnSts
   RUNG wire#powerrail
      Contact( #s150_ChkOprnSts )
      I_Contact( #sStWtResetRel )
      Contact( #sSst )
      wire#w1
      Contact( #c150_ChkOprnSts_T1 )
      Coil( #s150_ChkOprnSts_T1 )
   END_RUNG
   RUNG wire#w1
      I_Contact( #s150_ChkOprnSts_T1 )
      Contact( #c150_ChkOprnSts_T2 )
      Coil( #s150_ChkOprnSts_T2 )
   END_RUNG
   // the same network as SCL:
   #_w1 := #s150_ChkOprnSts AND NOT #sStWtResetRel AND #sSst;
   #s150_ChkOprnSts_T1 := #_w1 AND #c150_ChkOprnSts_T1;
   #s150_ChkOprnSts_T2 := #_w1 AND NOT #s150_ChkOprnSts_T1 AND #c150_ChkOprnSts_T2;
END_REGION

REGION Network 55: STATE Num:150 ChkOprnSts
   RUNG wire#powerrail
      Contact( #s150_ChkOprnSts )
      wire#w1
      I_Contact( #sStWtResetRel )
      I_Contact( #s150_ChkOprnSts_T1 )
      I_Contact( #s150_ChkOprnSts_T2 )
      wire#w2
      Coil( #s150_ChkOprnSts )
   END_RUNG
   RUNG wire#powerrail
      Contact( #s30_ChkPartPrsnt_T1 )
   END_RUNG wire#w1
   RUNG wire#w2
      { S7_GenerateENO := "TRUE" } Move(in := 150, out1 => #qStateNo)
   END_RUNG
   // the same network as SCL:
   #s150_ChkOprnSts := (#s150_ChkOprnSts OR #s30_ChkPartPrsnt_T1) AND NOT #sStWtResetRel AND NOT #s150_ChkOprnSts_T1 AND NOT #s150_ChkOprnSts_T2;
   IF #s150_ChkOprnSts THEN #qStateNo := 150; END_IF;
END_REGION
END_FUNCTION_BLOCK
